TYPE ST_HmiBrakeStatus :
STRUCT
	bPresent	: BOOL;
	bOpen		: BOOL;
END_STRUCT
END_TYPE

(* stored: Version 1.1.0.1, ProductVersion 3.1.4024.15
   DUT ST_HmiBrakeStatus: Id {687968ef-069b-45ca-917f-e30bc7eb7e64} *)
